TYPE ST_ControlModuleDevList :
STRUCT
	DiMomentaryPb	: I_DevDigitalIn;
	CylExample		: I_DevCylinder;
	DoSignalPl		: I_DevDigitalOut;
END_STRUCT
END_TYPE

(* stored: Version 1.1.0.1, ProductVersion 3.1.4024.12
   DUT ST_ControlModuleDevList: Id {478f85a9-c35e-49e7-a233-0395b519f793} *)
